(* IEC 61131-3 sources: JingjiangMoonbox/Application/Application/数据类型/通讯协议/子影, 5 files *)

(* ---- StParam_UnitHMI485_Rd.st ---- *)
(*@CES
Name=StParam_UnitHMI485_Rd
Type=Gvl
TypeGuid=2db5746d-d284-4425-9f7f-2663a34b0ebc
Guid=b1f3dc45-0cc5-41fd-a54e-f4937ddba804
HasDeclaration=True
HasImplementation=False
*)
{DECLARATION}
{attribute 'pack_mode' := '1'}
TYPE StParam_UnitHMI485_Rd :
STRUCT
//每个包240字节
//新增读取内容||工艺控制相关2025.12.31.135951||总共24字节||120-24=96
	rHz_UnitInkRoller_CurrRD: REAL;
	wSts_UnitInkRoller: WORD;
	rHz_UnitScraper_CurrRD: REAL;
	wSts_UnitScraper: WORD;
	rHz_UnitHotWind_CurrRd: REAL;
	wSts_UnitHotWind: WORD;
	rHz_UnitHotWind_CurrRd_2: REAL;
	wSts_UnitHotWind_2: WORD;

	abyRsv_Rd: ARRAY [1..96] OF BYTE;(*只读通讯保留位*)

//第二个人机通讯内容2025.12.31.154101
	rHz_UnitInkRoller_CurrRD_OtherUnit: REAL;
	wSts_UnitInkRoller_OtherUnit: WORD;
	rHz_UnitScraper_CurrRD_OtherUnit: REAL;
	wSts_UnitScraper_OtherUnit: WORD;
	rHz_UnitHotWind_CurrRd_OtherUnit: REAL;
	wSts_UnitHotWind_OtherUnit: WORD;
	rHz_UnitHotWind_CurrRd_2_OtherUnit: REAL;
	wSts_UnitHotWind_2_OtherUnit: WORD;
	abyRsv_Rd_OtherUnit: ARRAY [1..96] OF BYTE;(*只读通讯保留位*)

END_STRUCT
END_TYPE

{IMPLEMENTATION}

(* ---- StParam_UnitHMI485_Wr_81.st ---- *)
(*@CES
Name=StParam_UnitHMI485_Wr_81
Type=Gvl
TypeGuid=2db5746d-d284-4425-9f7f-2663a34b0ebc
Guid=7390c00c-e7d7-4035-8319-06dcd475a32f
HasDeclaration=True
HasImplementation=False
*)
{DECLARATION}
{attribute 'pack_mode' := '1'}
TYPE StParam_UnitHMI485_Wr_81 :
STRUCT
	byPackId: BYTE;//先放一个标志标记通讯只写内容的格式：
	//=1--StParam_UnitHMI485_Wr_81
	//=2--StParam_UnitHMI485_Wr_82
	//=3--StParam_UnitHMI485_Wr_83
	wGirth: WORD;(*版周长*10*)
	iCompanyId: INT;(*用户编号*)
	iPromptMsgId: INT;(*当前报警/提示信息*)
	wAxisId_And_GrpId: WORD;(*高8位轴号，低8位系号*)
	wLedtime_And_Language: WORD;(*高8位屏保延时，低8位语言选择*)
	aiErrorBuff_V: ARRAY [1..40] OF INT;(*纵向误差队列*)
	aiErrorBuff_H: ARRAY [1..40] OF INT;(*横向误差队列*)
	iVel_Axis: INT;(*轴速度*10*)
	iVel_Grp: INT;(*系速度*10*)
	wIndex_And_ErrNum: WORD;(*高8为采样索引，低8为误差刷新幅数*)
	iArcAlarm_V: INT;(*纵向报警值*)
	iArcAlarm_H: INT;(*横向报警值*)
	wFlag_Arc: WORD;(*套色相关标志，bit0-bit6:色标形式；bit7-bot11:色标顺逆序；bit12:压辊状态*)
	wLED_485Cnt: WORD;(*高8为屏保图片，低8为485通讯计数*)
	wUnit_Input_I: WORD;(*IO监控输入*)
	wUnit_Input_II: WORD;(*IO监控输入*)
	wUnit_Input_III: WORD;(*IO监控输入*)
	wHz_UnitInkRoller_CurrWR: WORD;(*递墨辊频率写入值*)
	wHz_UnitScraper_CurrWR: WORD;(*刮刀频率写入值*)
	wHz_UnitHotWind_CurrWR: WORD;(*热风频率写入值*)
	wHz_UnitHotWind2_CurrWR: WORD;(*热风频率写入值*)
	wPV_UnitTemCtl: WORD;(*实时温度*)
	wSts_UnitTemCtl: WORD;(*加热状态*)
	rPos_PrnRoller_Pressure_M							: REAL;(* 版辊压力电机位置M侧/实时值|mm-根据坐标系变化 *)
	rPos_PrnRoller_Pressure_G							: REAL;(* 版辊压力电机位置G侧/实时值|mm-根据坐标系变化 *)
	rPos_NetRoller_Pressure_M							: REAL;(* 网辊压力电机位置M侧/实时值|mm-根据坐标系变化 *)
	rPos_NetRoller_Pressure_G							: REAL;(* 网辊压力电机位置G侧/实时值|mm-根据坐标系变化 *)

	bySts_Ctl: BYTE;//留有一个BYTE作为通讯一些重要标志
	//BIT0:先用作第二色组通讯使能2026.1.4.140126
	abyRsv_HignComm: ARRAY [1..20] OF BYTE;(*保留24个寄存器*)

END_STRUCT
END_TYPE

{IMPLEMENTATION}

(* ---- StParam_UnitHMI485_Wr_82.st ---- *)
(*@CES
Name=StParam_UnitHMI485_Wr_82
Type=Gvl
TypeGuid=2db5746d-d284-4425-9f7f-2663a34b0ebc
Guid=726df55c-874d-4dcc-bc3a-20d650b779ca
HasDeclaration=True
HasImplementation=False
*)
{DECLARATION}
{attribute 'pack_mode' := '1'}
TYPE StParam_UnitHMI485_Wr_82 ://全部作为预留区域||2026.1.4.135806
STRUCT
	byPackId: BYTE;//先放一个标志标记通讯只写内容的格式：
	//=1--StParam_UnitHMI485_Wr_81
	//=2--StParam_UnitHMI485_Wr_82
	//=3--StParam_UnitHMI485_Wr_83
	abyRsv_LowComm: ARRAY [1..239] OF BYTE;(*低速只写通讯保留位*)
END_STRUCT
END_TYPE

{IMPLEMENTATION}

(* ---- StParam_UnitHMI485_Wr_83.st ---- *)
(*@CES
Name=StParam_UnitHMI485_Wr_83
Type=Gvl
TypeGuid=2db5746d-d284-4425-9f7f-2663a34b0ebc
Guid=f4069e2c-8ef0-4053-8cd1-9b1dedc27d09
HasDeclaration=True
HasImplementation=False
*)
{DECLARATION}
{attribute 'pack_mode' := '1'}
TYPE StParam_UnitHMI485_Wr_83 ://作为第二色组通讯内容2026.1.4.135901||在Wr-81里增加第二色组通讯使能
STRUCT
	byPackId: BYTE;//先放一个标志标记通讯只写内容的格式：
	//=1--StParam_UnitHMI485_Wr_81
	//=2--StParam_UnitHMI485_Wr_82
	//=3--StParam_UnitHMI485_Wr_83
	wGirth_OtherUnit: WORD;(*版周长*10*)
	iCompanyId_OtherUnit: INT;(*用户编号*)
	iPromptMsgId_OtherUnit: INT;(*当前报警/提示信息*)
	wAxisId_And_GrpId_OtherUnit: WORD;(*高8位轴号，低8位系号*)
	wLedtime_And_Language_OtherUnit: WORD;(*高8位屏保延时，低8位语言选择*)
	iVel_Axis_OtherUnit: INT;(*轴速度*10*)
	iVel_Grp_OtherUnit: INT;(*系速度*10*)
	wIndex_And_ErrNum_OtherUnit: WORD;(*高8为采样索引，低8为误差刷新幅数*)
	wFlag_Arc_OtherUnit: WORD;(*套色相关标志，bit0-bit6:色标形式；bit7-bot11:色标顺逆序；bit12:压辊状态*)
	wLED_485Cnt_OtherUnit: WORD;(*高8为屏保图片，低8为485通讯计数*)
	wUnit_Input_I_OtherUnit: WORD;(*IO监控输入*)
	wUnit_Input_II_OtherUnit: WORD;(*IO监控输入*)
	wUnit_Input_III_OtherUnit: WORD;(*IO监控输入*)
	wHz_UnitInkRoller_CurrWR_OtherUnit: WORD;(*递墨辊频率写入值*)
	wHz_UnitScraper_CurrWR_OtherUnit: WORD;(*刮刀频率写入值*)
	wHz_UnitHotWind_CurrWR_OtherUnit: WORD;(*热风频率写入值*)
	wHz_UnitHotWind2_CurrWR_OtherUnit: WORD;(*热风频率写入值*)
	wPV_UnitTemCtl_OtherUnit: WORD;(*实时温度*)
	wSts_UnitTemCtl_OtherUnit: WORD;(*加热状态*)
	rPos_PrnRoller_Pressure_M_OtherUnit							: REAL;(* 版辊压力电机位置M侧/实时值|mm-根据坐标系变化 *)
	rPos_PrnRoller_Pressure_G_OtherUnit							: REAL;(* 版辊压力电机位置G侧/实时值|mm-根据坐标系变化 *)
	rPos_NetRoller_Pressure_M_OtherUnit							: REAL;(* 网辊压力电机位置M侧/实时值|mm-根据坐标系变化 *)
	rPos_NetRoller_Pressure_G_OtherUnit							: REAL;(* 网辊压力电机位置G侧/实时值|mm-根据坐标系变化 *)

	abyRsv_HignComm_OtherUnit: ARRAY [1..185] OF BYTE;(*保留120个寄存器*)
//2025.11.27.181845增加压力相关内容占用 64字节，剩余字节120-64=56
//	awRsv_HignComm_2: ARRAY [1..120] OF WORD;(*保留120个寄存器*)
END_STRUCT
END_TYPE

{IMPLEMENTATION}

(* ---- StParam_UnitHMI485_WrRd.st ---- *)
(*@CES
Name=StParam_UnitHMI485_WrRd
Type=Gvl
TypeGuid=2db5746d-d284-4425-9f7f-2663a34b0ebc
Guid=20b40184-5295-49e6-bf5f-17e6b491675e
HasDeclaration=True
HasImplementation=False
*)
{DECLARATION}
{attribute 'pack_mode' := '1'}
TYPE StParam_UnitHMI485_WrRd :
STRUCT
	byHMI_Cnt: BYTE;(*人机通讯计数*)
	byAxisId: BYTE;(*轴号*)
	iAdjust_V: INT;(*套色修正量，单位：丝*)
	iAdjust_H: INT;(*套色修正量，单位：丝*)
	wStatus: WORD;(*界面上套色相关状态*)
	wButtonFun: WORD;(*界面按钮及指示灯*)
	wSwitchFun: WORD;(*界面开关*)
	wUnit_Outout_I: WORD;(*IO输出监控/测试*)
	wUnit_Outout_II: WORD;(*IO输出监控/测试*)
	iPlateAdjustmentProf:INT;(*纵向快速对版量*)
	iJourney_HorzRapidAdjust: INT;(*横向快速对版量*)
	wHz_UnitInkRoller_ManuallySet: WORD;(*递墨辊手动频率*)
	wCoeff_UnitInkRoller_Auto: WORD;(*递墨辊自动系数*)
	wHz_UnitScraper_ManuallySet: WORD;(*刮刀手动频率*)
	wCoeff_UnitScraper_Auto: WORD;(*刮刀自动系数*)
	wHz_UnitHotWind: WORD;(*热风频率*)
	wHz_UnitHotWind_2: WORD;(*热风2频率*)
	wSV_UnitTemCtl: WORD;(*加热设定温度*)
	dwCtlBits_UnitBaseCraft: DWORD;(*工艺控制开关*)
	wAirInletWindDoorValue: WORD;(*进风风门*)
	wAirExhaustWindDoorValue: WORD;(*排风风门*)
	wAirReturnWindDoorValue: WORD;(*回风风门*)
//增加一些开关变量||2025.12.31.141711||总共	7||94-7=87
	bySwitch_Arc: BYTE;(*先用一个BYTE作为其他套色需要的开关
							bit0: 横向开关*)
	wSwitch_Process: WORD;(*工艺开关
							bit0:递墨辊自动
							bit1:递墨辊正转
							bit2:递墨辊反转
							bit3:刮刀自动
							bit4:刮刀开关
							bit5:加热I档
							bit6:加热II档
							bit7:加热III档
							bit8:热风开关
							bit9:热风2开关
*)
	dwSwitch_Pressure: DWORD;(*压力相关
							bit0:版辊压力操作侧靠近
							bit1:版辊压力操作侧远离
							bit2:版辊压力传动侧靠近
							bit3:版辊压力传动侧远离
							bit4:版辊压力靠近
							bit5:版辊压力远离
							bit6:网辊压力操作侧靠近
							bit7:网辊压力操作侧远离
							bit8:网辊压力传动侧靠近
							bit9:网辊压力传动侧远离
							bit10:网辊压力靠近
							bit11:网辊压力远离
							bit12:张带辊压力操作侧靠近
							bit13:张带辊压力操作侧远离
							bit14:张带辊压力传动侧靠近
							bit15:张带辊压力传动侧远离
							bit16:张带辊压力靠近
							bit17:张带辊压力远离
							bit18~bit23:预留
							bit24:版辊离压位标定
							bit25:版辊合压位标定
							bit26:版辊换版位标定
							bit27:版辊平行标定
							bit24:网辊离压位标定
							bit25:网辊合压位标定
							bit26:网辊换版位标定
							bit27:网辊平行标定
*)
	abyRsv_RdWr: ARRAY [1..73] OF BYTE;

	byHMI_Cnt_OtherUnit: BYTE;(*人机通讯计数*)
	byAxisId_OtherUnit: BYTE;(*轴号*)
	wButtonFun_OtherUnit: WORD;(*界面按钮及指示灯*)
	wSwitchFun_OtherUnit: WORD;(*界面开关*)
	wUnit_Outout_I_OtherUnit: WORD;(*IO输出监控/测试*)
	wUnit_Outout_II_OtherUnit: WORD;(*IO输出监控/测试*)
	iJourney_HorzRapidAdjust_OtherUnit: INT;(*横向快速对版量*)
	wHz_UnitInkRoller_ManuallySet_OtherUnit: WORD;(*递墨辊手动频率*)
	wCoeff_UnitInkRoller_Auto_OtherUnit: WORD;(*递墨辊自动系数*)
	wHz_UnitScraper_ManuallySet_OtherUnit: WORD;(*刮刀手动频率*)
	wCoeff_UnitScraper_Auto_OtherUnit: WORD;(*刮刀自动系数*)
	wHz_UnitHotWind_OtherUnit: WORD;(*热风频率*)
	wHz_UnitHotWind_2_OtherUnit: WORD;(*热风2频率*)
	wSV_UnitTemCtl_OtherUnit: WORD;(*加热设定温度*)
	dwCtlBits_UnitBaseCraft_OtherUnit: DWORD;(*工艺控制开关*)
	wAirInletWindDoorValue_OtherUnit: WORD;(*进风风门*)
	wAirExhaustWindDoorValue_OtherUnit: WORD;(*排风风门*)
	wAirReturnWindDoorValue_OtherUnit: WORD;(*回风风门*)
//增加一些开关变量||2025.12.31.141711||总共	7||94-7=87
	wSwitch_Process_OtherUnit: WORD;(*工艺开关
							bit0:递墨辊自动
							bit1:递墨辊正转
							bit2:递墨辊反转
							bit3:刮刀自动
							bit4:刮刀开关
							bit5:加热I档
							bit6:加热II档
							bit7:加热III档
							bit8:热风开关
							bit9:热风2开关
*)
	dwSwitch_Pressure_OtherUnit: DWORD;(*压力相关
							bit0:版辊压力操作侧靠近
							bit1:版辊压力操作侧远离
							bit2:版辊压力传动侧靠近
							bit3:版辊压力传动侧远离
							bit4:版辊压力靠近
							bit5:版辊压力远离
							bit6:网辊压力操作侧靠近
							bit7:网辊压力操作侧远离
							bit8:网辊压力传动侧靠近
							bit9:网辊压力传动侧远离
							bit10:网辊压力靠近
							bit11:网辊压力远离
							bit12:张带辊压力操作侧靠近
							bit13:张带辊压力操作侧远离
							bit14:张带辊压力传动侧靠近
							bit15:张带辊压力传动侧远离
							bit16:张带辊压力靠近
							bit17:张带辊压力远离
							bit18~bit23:预留
							bit24:版辊离压位标定
							bit25:版辊合压位标定
							bit26:版辊换版位标定
							bit27:版辊平行标定
							bit24:网辊离压位标定
							bit25:网辊合压位标定
							bit26:网辊换版位标定
							bit27:网辊平行标定
*)
	abyRsv_RdWr_OtherUnit: ARRAY [1..74] OF BYTE;

END_STRUCT
END_TYPE

{IMPLEMENTATION}
